Staubli VAL3: Lab2A_L3.dtx


